// The only PLC data the HMI uses. Both structs are mapped automatically into
// the TwinCAT HMI server (attribute TcHmiSymbol.AddSymbol).
{attribute 'qualified_only'}
VAR_GLOBAL
    {attribute 'TcHmiSymbol.AddSymbol'}
    stStatus  : ST_HmiStatus;
    {attribute 'TcHmiSymbol.AddSymbol'}
    stCommand : ST_HmiCommand;
END_VAR

(* stored: Version 1.1.0.1
   GVL GVL_Hmi: Id {56ec23f2-91ad-16cb-49e7-68d04d488fac} *)
